FUNCTION_BLOCK DLG_Toast (* Hinweis ohne Tasten, verschwindet nach TIMEOUT *)
  (* Standard: 61499-2; Description: Copyright (c) 2026 Meisterschulen am Ostbahnhof This program and the accompanying materials are made available under the terms of the Eclipse Public License 2.0 which is available at https://www.eclipse.org/legal/epl-2.0/ SPDX-License-Identifier: EPL-2.0 *)
  (* Version 1.1, 2026-11-25, Franz Höpfinger, Meisterschulen am Ostbahnhof, SubApp -> Composite FB (Lib wird wegen DLG_CTRL ohnehin gebaut, im fboot nur eine Instanz). *)
  (* Version 1.0, 2026-11-17, Franz Höpfinger, Meisterschulen am Ostbahnhof, initial API and implementation and/or initial documentation *)
  PACKAGE isobus::UT::dialog;
  IMPORT isobus::UT::Q::const::IDs::ID_NULL;
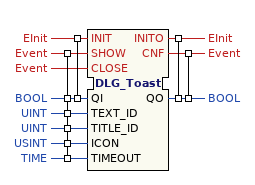
  EVENT_INPUT
    INIT : EInit WITH QI; (* Initialisierung *)
    SHOW WITH QI, TEXT_ID, TITLE_ID, ICON, TIMEOUT; (* Hinweis zeigen *)
    CLOSE; (* Hinweis schliessen *)
  END_EVENT
  EVENT_OUTPUT
    INITO : EInit WITH QO; (* Initialisierung fertig *)
    CNF WITH QO; (* Hinweis beendet *)
  END_EVENT
  VAR_INPUT
    QI : BOOL := TRUE; (* Freigabe *)
    TEXT_ID : UINT := ID_NULL; (* OutputString Meldungstext *)
    TITLE_ID : UINT := ID_NULL; (* OutputString Titel, NULL = Standard *)
    ICON : USINT := USINT#1; (* DLG_ICON_* *)
    TIMEOUT : TIME := T#3s; (* Anzeigedauer *)
  END_VAR
  VAR_OUTPUT
    QO : BOOL; (* Qualitaet *)
  END_VAR
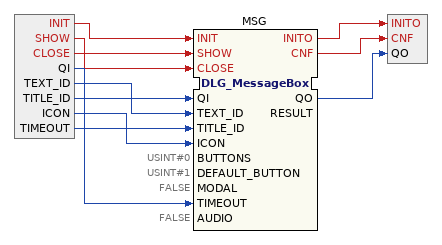
  FBS
    MSG : isobus::UT::dialog::DLG_MessageBox(BUTTONS := USINT#0, DEFAULT_BUTTON := USINT#1, MODAL := FALSE, AUDIO := FALSE);
  END_FBS
  EVENT_CONNECTIONS
    INIT TO MSG.INIT;
    MSG.INITO TO INITO;
    SHOW TO MSG.SHOW;
    CLOSE TO MSG.CLOSE;
    MSG.CNF TO CNF;
  END_CONNECTIONS
  DATA_CONNECTIONS
    QI TO MSG.QI;
    TEXT_ID TO MSG.TEXT_ID;
    TITLE_ID TO MSG.TITLE_ID;
    ICON TO MSG.ICON;
    TIMEOUT TO MSG.TIMEOUT;
    MSG.QO TO QO;
  END_CONNECTIONS
END_FUNCTION_BLOCK
